{region 'Documentation'}
(*!
<summary>Checks that the falling-edge count is inside the inclusive range.</summary>
<description>

Reversed bounds report Error during evaluation; equal bounds are valid.

Observation and accumulated-count handling come from AssertionEdgeCountBase. Evaluate
checks the held count independently of Enable; reset clears the count and baseline.

</description>
*)
{endregion}
FUNCTION_BLOCK AssertFallingEdgeCntInRange EXTENDS AssertionEdgeCountBase
VAR_INPUT
    Minimum : UINT; //! Inclusive lower bound of the comparison; for a range, must not exceed Maximum.
    Maximum : UINT; //! Inclusive upper bound of the comparison; for a range, must not be below Minimum.
END_VAR

SUPER^();

{region 'Documentation'}
(*!
<summary>Observe through the base, then evaluate the count with Error priority.</summary>
*)
{endregion}
METHOD PROTECTED Assert
VAR
    Message : STRING(GVL_Constants.MessageLength);
    MinimumText : STRING(GVL_Constants.AssertionValueLength);
    MaximumText : STRING(GVL_Constants.AssertionValueLength);
    ActualText : STRING(GVL_Constants.AssertionValueLength);
END_VAR
SUPER^.Assert();

IF NOT EvaluationActive THEN
    RETURN;
END_IF;

IF Result = E_Result.Error THEN
    RETURN;
END_IF;

IF Minimum > Maximum THEN
    MinimumText := UINT_TO_STRING(Minimum);
    MaximumText := UINT_TO_STRING(Maximum);
    Message := CONCAT('Assertion error: minimum exceeds maximum. Minimum = ',
        MinimumText);
    Message := CONCAT(Message, ', Maximum = ');
    Message := CONCAT(Message, MaximumText);
    Message := CONCAT(Message, '.');
    Error(Message := Message);
    RETURN;
END_IF;

IF Result = E_Result.Failed THEN
    RETURN;
END_IF;

IF (EdgeCount < Minimum) OR (EdgeCount > Maximum) THEN
    MinimumText := UINT_TO_STRING(Minimum);
    MaximumText := UINT_TO_STRING(Maximum);
    ActualText := UINT_TO_STRING(EdgeCount);
    Message := CONCAT('Assertion failed: falling edge count is outside allowed range. Minimum = ',
        MinimumText);
    Message := CONCAT(Message, ', Maximum = ');
    Message := CONCAT(Message, MaximumText);
    Message := CONCAT(Message, ', Actual = ');
    Message := CONCAT(Message, ActualText);
    Message := CONCAT(Message, '.');
    Fail(Message := Message);
    RETURN;
END_IF;

Pass();
END_METHOD

{region 'Documentation'}
(*!
<summary>Recognize a falling edge without changing observation state.</summary>
*)
{endregion}
METHOD PROTECTED IsMatchingEdge : BOOL //! TRUE when PreviousValue and CurrentValue form the edge selected by this Assertion.
VAR_INPUT
    PreviousValue : BOOL; //! Signal value from the preceding active observation.
    CurrentValue : BOOL; //! Signal value from the current active observation.
END_VAR
IsMatchingEdge := PreviousValue AND NOT CurrentValue;
END_METHOD

END_FUNCTION_BLOCK

(* stored: Version 1.1.0.1
   POU AssertFallingEdgeCntInRange: Id {14bdcc68-396f-48bf-b27c-caf4aff98a64}, SpecialFunc None
   Folder Internal: Id {960b0c65-daa7-4266-8a43-701cee310969}
   Method Assert: Id {aa4fac57-5741-45bf-9c2c-fa92ea1805bd}
   Method IsMatchingEdge: Id {b2f05f1a-b42a-409c-a90b-dc3c11007381} *)
